// TIA Portal project "Conveyor_Control_V17" (V17)
// Vorlageprojekt für das Buch mit Zielsystem S7-1200

(* hardware
DEVICE "S7-1200-Station_1"  S7-1200 Station
   slot 0: "Baugruppenträger_0"  Rack  V1.0
   slot 1: "PLC_1"  CPU 1211C DC/DC/DC  6ES7 211-1AE40-0XB0  V4.1
*)

// ===== PLC "PLC_1"  CPU 1211C DC/DC/DC =====

VAR_GLOBAL   // PLC tag table "Standard-Variablentabelle"
   "PB_Start" AT %I0.0 : Bool;
   "PB_Stop" AT %I0.1 : Bool;
   "Mode_Auto" AT %I0.2 : Bool;
   "Mode_Manual" AT %I0.3 : Bool;
   "Manual_Jog" AT %I0.4 : Bool;
   "Sensor_Product" AT %I0.5 : Bool;
   "PB_Reset" AT %I0.6 : Bool;
   "Falla_Simulada" AT %I0.7 : Bool;
   "Motor_Conveyor" AT %Q0.0 : Bool;
   "Lamp_Run" AT %Q0.1 : Bool;
   "Lamp_Fault" AT %Q0.2 : Bool;
   "Lamp_Done" AT %Q0.3 : Bool;
END_VAR

// folder: Conveyor

DATA_BLOCK "Variables"   // DB1
{ S7_Optimized_Access := 'TRUE' }
VERSION : 0.1
   VAR
      Permissie_Ok : Bool;   // Permiso de funcionamiento
      Auto_Run_Latch : Bool;   // Memoria de ciclo Automatico
      Manual_Run_Cmd : Bool;   // Solcitud de marcha Manual
      Motor_Run_Cmd_1 : Bool;   // Comando logico final
      Product_Pulse : Bool;   // Pulso de un solo ciclo por deteccion
      Cycle_Done : Bool;   // Objetivo de produccion alcanzado
      Product_Count : Int;   // Cantidad de productos detectados
      Step_Machine : Int;
   END_VAR
BEGIN
END_DATA_BLOCK

// folder: System blocks/Program resources

DATA_BLOCK "CTU_Procuction"   // DB3
{ S7_Optimized_Access := 'TRUE' }
AUTHOR : Simatic
FAMILY : IEC
NAME : CNTR
VERSION : 1.0
// stored: InstanceOfName IEC_COUNTER
"IEC_COUNTER"
BEGIN
END_DATA_BLOCK

// folder: (top level)

FUNCTION "MHJ-PLC-Lab-Function-S71200" : Void   // FC9000, SCL
{ S7_Optimized_Access := 'TRUE' }
VERSION : 0.1
   VAR_TEMP
      rdTimeReturn : Int;
      outputTime : DTL;
      SyncVal : Byte;
      forVal : Int;
      forVal_2 : Int;
      Value : Byte;
   END_VAR
   VAR CONSTANT
      CompVal : Byte := 16#34;
      Value_01 : Byte := 16#11;
      Value_01_DW : DWord := 16#A165_D992;
      Value_02_DW : DWord := 16#58BE_4401;
   END_VAR
BEGIN

   #Value:=PEEK(area := 16#82,
        dbNumber := 0,
        byteOffset := 511);
   #Value := #Value + 1;

   POKE(area := 16#82,
        dbNumber := 0,
        byteOffset := 511,
        value := #Value);

   POKE(area:=16#81,
        dbNumber:=0,
        byteOffset:=1016,
        value:=#Value_01_DW);
   POKE(area := 16#81,
        dbNumber := 0,
        byteOffset := 1020,
        value := #Value_02_DW);

   POKE(area := 16#81,
        dbNumber := 0,
        byteOffset := 511,
        value := B#16#00);

   FOR #forVal := 0 TO 120 DO
       FOR #forVal_2:=0 TO 10 DO
           #rdTimeReturn:=RD_SYS_T(#outputTime);
           #rdTimeReturn := WR_SYS_T(#outputTime);
           #rdTimeReturn := RD_SYS_T(#outputTime);
           #rdTimeReturn := WR_SYS_T(#outputTime);
       END_FOR;
       #SyncVal:= PEEK(area := 16#81,
                      dbNumber := 0,
                      byteOffset := 511);
       IF #SyncVal = #CompVal THEN
          GOTO M_1;
       END_IF;
   END_FOR;
   RETURN;

   M_1:
   POKE(area := 16#81,
        dbNumber := 0,
        byteOffset := 511,
        value := B#16#0);
END_FUNCTION

ORGANIZATION_BLOCK "Main"   // OB1, FBD, ProgramCycle
TITLE = "Main Program Sweep (Cycle)"
{ S7_Optimized_Access := 'TRUE' }
VERSION : 0.1
   VAR_INPUT
      Initial_Call : Bool;   // Initial call of this OB
      Remanence : Bool;   // =True, if remanent data are available
   END_VAR
   VAR_TEMP   // added for the SCL form of the ladder/FBD networks
      _w1 : Bool;
   END_VAR
BEGIN

REGION Network 1: Konnektierungsbaustein für PLC-Lab
   // Im Netzwerk 1 wird der Konnektierungsbaustein für PLC-Lab aufgerufen.
   // Dieser Aufruf darf nicht entfernt werden!
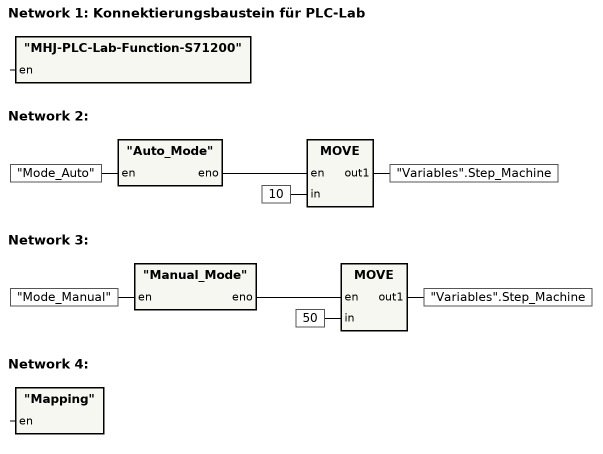
   "MHJ-PLC-Lab-Function-S71200"();
END_REGION

REGION Network 2
   // AutoMode
   "Auto_Mode"(EN := "Mode_Auto", ENO => #_w1);
   IF #_w1 THEN "Variables".Step_Machine := 10; END_IF;
END_REGION

REGION Network 3
   // ManualMode
   "Manual_Mode"(EN := "Mode_Manual", ENO => #_w1);
   IF #_w1 THEN "Variables".Step_Machine := 50; END_IF;
END_REGION

REGION Network 4
   "Mapping"();
END_REGION
END_ORGANIZATION_BLOCK

// folder: Conveyor

FUNCTION "Auto_Mode" : Void   // FC1, LAD
{ S7_Optimized_Access := 'TRUE' }
VERSION : 0.1
   VAR_TEMP   // added for the SCL form of the ladder/FBD networks
      _w1 : Bool;
   END_VAR
BEGIN

REGION Network 1: Permiso de funcionamiento
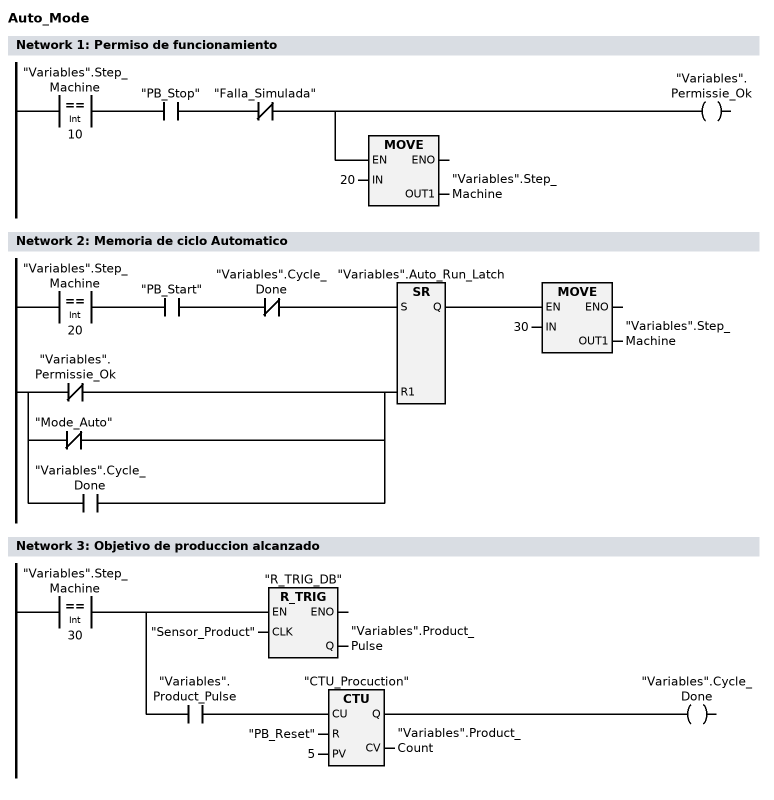
   RUNG wire#powerrail
      { S7_Templates := "SrcType := Int" } EQ_Contact(in1 := "Variables".Step_Machine, in2 := 10)
      Contact( "PB_Stop" )
      I_Contact( "Falla_Simulada" )
      wire#w1
      Coil( "Variables".Permissie_Ok )
   END_RUNG
   RUNG wire#w1
      Move(in := 20, out1 => "Variables".Step_Machine)
   END_RUNG
   // the same network as SCL:
   "Variables".Permissie_Ok := ("Variables".Step_Machine = 10) AND "PB_Stop" AND NOT "Falla_Simulada";
   IF "Variables".Permissie_Ok THEN "Variables".Step_Machine := 20; END_IF;
END_REGION

REGION Network 2: Memoria de ciclo Automatico
   RUNG wire#powerrail
      { S7_Templates := "SrcType := Int" } EQ_Contact(in1 := "Variables".Step_Machine, in2 := 20)
      Contact( "PB_Start" )
      I_Contact( "Variables".Cycle_Done )
      S_SR(operand := "Variables".Auto_Run_Latch, r1 := wire#w1)
      Move(in := 30, out1 => "Variables".Step_Machine)
   END_RUNG
   RUNG wire#powerrail
      I_Contact( "Variables".Permissie_Ok )
   END_RUNG wire#w1
   RUNG wire#powerrail
      I_Contact( "Mode_Auto" )
   END_RUNG wire#w1
   RUNG wire#powerrail
      Contact( "Variables".Cycle_Done )
   END_RUNG wire#w1
   // the same network as SCL:
   IF ("Variables".Step_Machine = 20) AND "PB_Start" AND NOT "Variables".Cycle_Done THEN
       "Variables".Auto_Run_Latch := TRUE;   // SR flip-flop
   END_IF;
   IF NOT "Variables".Permissie_Ok OR NOT "Mode_Auto" OR "Variables".Cycle_Done THEN
       "Variables".Auto_Run_Latch := FALSE;
   END_IF;
   IF "Variables".Auto_Run_Latch THEN "Variables".Step_Machine := 30; END_IF;
END_REGION

REGION Network 3: Objetivo de produccion alcanzado
   #_w1 := "Variables".Step_Machine = 30;
   IF #_w1 THEN
       "R_TRIG_DB"(CLK := "Sensor_Product", Q => "Variables".Product_Pulse);   // R_TRIG
   END_IF;
   "CTU_Procuction".CTU(CU := #_w1 AND "Variables".Product_Pulse,
                        R := "PB_Reset",
                        PV := 5,
                        CV => "Variables".Product_Count);
   "Variables".Cycle_Done := "CTU_Procuction".Q;
END_REGION
END_FUNCTION

FUNCTION "Manual_Mode" : Void   // FC2, LAD
{ S7_Optimized_Access := 'TRUE' }
VERSION : 0.1
BEGIN

REGION Network 1: Permiso de funcionamiento
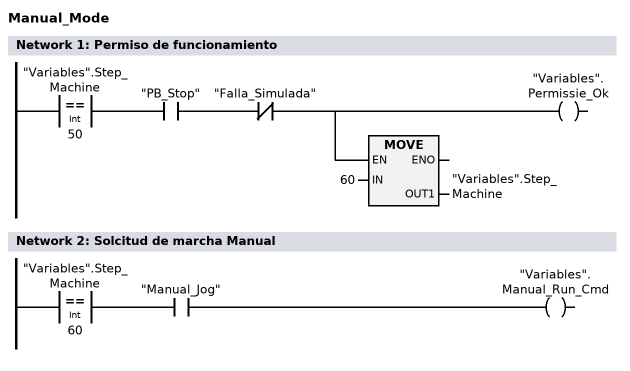
   RUNG wire#powerrail
      { S7_Templates := "SrcType := Int" } EQ_Contact(in1 := "Variables".Step_Machine, in2 := 50)
      Contact( "PB_Stop" )
      I_Contact( "Falla_Simulada" )
      wire#w1
      Coil( "Variables".Permissie_Ok )
   END_RUNG
   RUNG wire#w1
      Move(in := 60, out1 => "Variables".Step_Machine)
   END_RUNG
   // the same network as SCL:
   "Variables".Permissie_Ok := ("Variables".Step_Machine = 50) AND "PB_Stop" AND NOT "Falla_Simulada";
   IF "Variables".Permissie_Ok THEN "Variables".Step_Machine := 60; END_IF;
END_REGION

REGION Network 2: Solcitud de marcha Manual
   RUNG wire#powerrail
      { S7_Templates := "SrcType := Int" } EQ_Contact(in1 := "Variables".Step_Machine, in2 := 60)
      Contact( "Manual_Jog" )
      Coil( "Variables".Manual_Run_Cmd )
   END_RUNG
   // the same network as SCL:
   "Variables".Manual_Run_Cmd := ("Variables".Step_Machine = 60) AND "Manual_Jog";
END_REGION
END_FUNCTION

FUNCTION "Mapping" : Void   // FC3, LAD
{ S7_Optimized_Access := 'TRUE' }
VERSION : 0.1
BEGIN

REGION Network 1: Activacion de conveyor
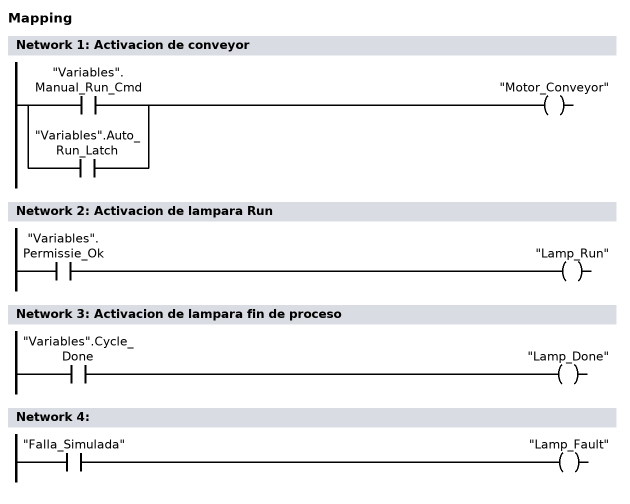
   RUNG wire#powerrail
      Contact( "Variables".Manual_Run_Cmd )
      wire#w1
      Coil( "Motor_Conveyor" )
   END_RUNG
   RUNG wire#powerrail
      Contact( "Variables".Auto_Run_Latch )
   END_RUNG wire#w1
   // the same network as SCL:
   "Motor_Conveyor" := "Variables".Manual_Run_Cmd OR "Variables".Auto_Run_Latch;
END_REGION

REGION Network 2: Activacion de lampara Run
   RUNG wire#powerrail
      Contact( "Variables".Permissie_Ok )
      Coil( "Lamp_Run" )
   END_RUNG
   // the same network as SCL:
   "Lamp_Run" := "Variables".Permissie_Ok;
END_REGION

REGION Network 3: Activacion de lampara fin de proceso
   RUNG wire#powerrail
      Contact( "Variables".Cycle_Done )
      Coil( "Lamp_Done" )
   END_RUNG
   // the same network as SCL:
   "Lamp_Done" := "Variables".Cycle_Done;
END_REGION

REGION Network 4
   RUNG wire#powerrail
      Contact( "Falla_Simulada" )
      Coil( "Lamp_Fault" )
   END_RUNG
   // the same network as SCL:
   "Lamp_Fault" := "Falla_Simulada";
END_REGION

REGION Network 5: Activacion de lampara de Falla
END_REGION
END_FUNCTION